(* IEC 61131-3 sources: PLC-Static-Analysis/modules/plc-rules/src/test/resources/PLCA-Q008, 2 files *)

(* ---- noncompliant.st ---- *)
PROGRAM P_Main
VAR
    fbMotor : FB_Motor;
    nCount : INT;
END_VAR
fbMotor();
nCount := F_Used(nCount);
END_PROGRAM

FUNCTION_BLOCK FB_Motor EXTENDS FB_Base
VAR
    bRun : BOOL;
END_VAR
bRun := NOT bRun;
END_FUNCTION_BLOCK

FUNCTION_BLOCK FB_Base
END_FUNCTION_BLOCK

FUNCTION_BLOCK FB_InGvl
END_FUNCTION_BLOCK

VAR_GLOBAL
    gfbSpare : FB_InGvl;
END_VAR

FUNCTION F_Used : INT
VAR_INPUT
    n : INT;
END_VAR
F_Used := F_Helper(n);
END_FUNCTION

FUNCTION F_Helper : INT
VAR_INPUT
    n : INT;
END_VAR
F_Helper := n + 1;
END_FUNCTION

FUNCTION F_Forgotten : INT // PLCA-Q008
VAR_INPUT
    n : INT;
END_VAR
F_Forgotten := F_Helper(n);
END_FUNCTION

FUNCTION_BLOCK FB_Old // PLCA-Q008
VAR
    n : INT;
END_VAR
n := 1;
END_FUNCTION_BLOCK

CONFIGURATION Cfg
    RESOURCE Res ON PLC
        TASK tMain(INTERVAL := T#10MS, PRIORITY := 1);
        PROGRAM iMain WITH tMain : P_Main;
    END_RESOURCE
END_CONFIGURATION

(* ---- compliant.st ---- *)
PROGRAM P_Main2
VAR
    nCount : INT;
END_VAR
nCount := F_Used2(nCount);
END_PROGRAM

FUNCTION F_Used2 : INT
VAR_INPUT
    n : INT;
END_VAR
F_Used2 := n + 1;
END_FUNCTION

CONFIGURATION Cfg2
    RESOURCE Res2 ON PLC
        TASK tMain2(INTERVAL := T#10MS, PRIORITY := 1);
        PROGRAM iMain2 WITH tMain2 : P_Main2;
    END_RESOURCE
END_CONFIGURATION
